{region 'Documentation'}
(*!
<summary>Checks that IN is NaN.</summary>
<description>

NaN and either infinity are legitimate checked data, not configuration errors.
Classification mismatch reports Failed. Bit-based classification does not perform an ordered
floating-point comparison.

Numeric diagnostics use the formatter's default six significant digits; rounding affects
the message only, not the comparison.

</description>
*)
{endregion}
FUNCTION_BLOCK AssertIsNaN_Real EXTENDS AssertionBase
VAR_INPUT
    IN : REAL; //! Value to classify; NaN and both infinities are valid inputs.
END_VAR

SUPER^();

{region 'Documentation'}
(*!
<summary>Classifies the bit representation without floating-point arithmetic.</summary>
*)
{endregion}
METHOD PROTECTED Assert
VAR
    Representation : AssertionRealRepresentation;
    Message : STRING(GVL_Constants.MessageLength);
END_VAR
VAR CONSTANT
    ExponentMask : DWORD := DWORD#16#7F800000;
    FractionMask : DWORD := DWORD#16#007FFFFF;
END_VAR
IF NOT EvaluationActive THEN
    RETURN;
END_IF;

IF Result = E_Result.Error THEN
    RETURN;
END_IF;

IF Result = E_Result.Failed THEN
    RETURN;
END_IF;

Representation.Value := IN;
IF ((Representation.Bits AND ExponentMask) <> ExponentMask)
    OR ((Representation.Bits AND FractionMask) = 0) THEN
    Message := CONCAT('Assertion failed: expected NaN. Actual = ',
        CreateAssertionTextValue_Real(Value := IN));
    Message := CONCAT(Message, '.');
    Fail(Message := Message);
    RETURN;
END_IF;

Pass();
END_METHOD

END_FUNCTION_BLOCK

(* stored: Version 1.1.0.1
   POU AssertIsNaN_Real: Id {d19d05de-1a00-4406-a637-7831b7984868}, SpecialFunc None
   Folder Internal: Id {9079145a-1988-4ebd-9da1-5280af06ad25}
   Method Assert: Id {a6310000-0000-4000-8000-000000000000} *)
